FUNCTION_BLOCK Actuator2OpBase (* Composite Function Block Type *)
  (* Standard: 61499-2 *)
  (* Version 1.0.1, 9/20/2023, ApplicationLibDevTeam, Schneider Electric, First Version *)
  PACKAGE Flexbridge.FestoMPS400;
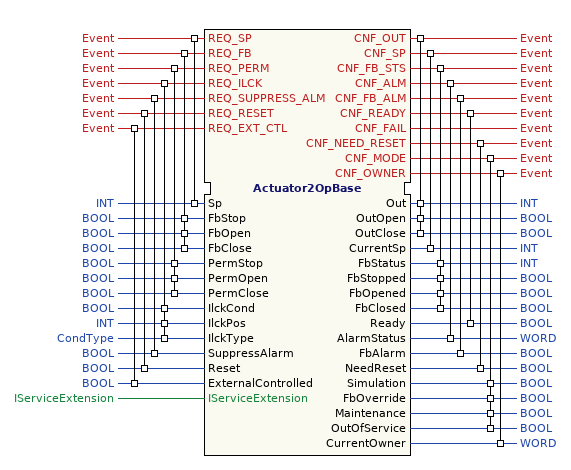
  EVENT_INPUT
    REQ_SP WITH Sp; (* Request to update setpoint *)
    REQ_FB WITH FbStop, FbOpen, FbClose; (* Request to update feedbacks *)
    REQ_PERM WITH PermStop, PermOpen, PermClose; (* Request to update permissive conditions *)
    REQ_ILCK WITH IlckCond, IlckPos, IlckType; (* Request to update interlock conditions *)
    REQ_SUPPRESS_ALM WITH SuppressAlarm; (* Request to update the alarm suppress status *)
    REQ_RESET WITH Reset; (* Request to reset the device *)
    REQ_EXT_CTL WITH ExternalControlled;
  END_EVENT
  EVENT_OUTPUT
    CNF_OUT WITH OutOpen, OutClose, Out; (* Execution confirmation of output *)
    CNF_SP WITH CurrentSp; (* Execution of confirmation Current Setpoint *)
    CNF_FB_STS WITH FbStopped, FbClosed, FbOpened, FbStatus; (* Execution of confirmed state *)
    CNF_ALM WITH AlarmStatus; (* Execution confirmation of alarm conditions *)
    CNF_FB_ALM WITH FbAlarm; (* Execution of confirmation  Fb alarm *)
    CNF_READY WITH Ready; (* Execution of Ready status *)
    CNF_FAIL; (* Execution of confirmation  failure *)
    CNF_NEED_RESET WITH NeedReset; (* Confirmation for resetting required *)
    CNF_MODE WITH Simulation, FbOverride, OutOfService, Maintenance; (* Excecution of new operational modes *)
    CNF_OWNER WITH CurrentOwner; (* Execution confirmation of owner *)
  END_EVENT
  VAR_INPUT
    Sp : INT; (* Setpoint of device (0 = Stop, 1 = Open, 2 =Close) *)
    FbStop : BOOL; (* 1 = Device stopfeedback active *)
    FbOpen : BOOL; (* 1 = Device open feedback active *)
    FbClose : BOOL; (* 1 = Device closed feedback active *)
    PermStop : BOOL := TRUE; (* 1 = Device stop permission active *)
    PermOpen : BOOL := TRUE; (* 1 = Device open permission active *)
    PermClose : BOOL := TRUE; (* 1 = Device close permission active *)
    IlckCond : BOOL; (* 1 = Interlock condition active *)
    IlckPos : INT; (* Interlock setpoint state (0 = Passive, 1 = Active1, 2 = Active2, 3 = Interlock inactive) *)
    IlckType : CondType; (* Type of condition interlock, (0 = Normal, 1 = Process interlock/Sequence interlock) *)
    SuppressAlarm : BOOL; (* 1 = Suppress alarm in HMI *)
    Reset : BOOL; (* 1 = Reset device failure *)
    ExternalControlled : BOOL; (* 1 = External control is active *)
  END_VAR
  VAR_OUTPUT
    Out : INT; (* Calculate output of the device ( 0 = Stop command, 1 = Open Command, 2 = Close Command) *)
    OutOpen : BOOL; (* 1 = Valve Output is Open *)
    OutClose : BOOL; (* 1 = Valve Output is Closed *)
    CurrentSp : INT; (* Output value considering permissive conditions *)
    FbStatus : INT; (* Confirmed state of the device (0 = Stopped, 1 = Opened, 2 = Closed,  253 = Unknown) *)
    FbStopped : BOOL; (* 1 = Stopped *)
    FbOpened : BOOL; (* 1 = Valve Open *)
    FbClosed : BOOL; (* 1 = Valve Closed *)
    Ready : BOOL; (* 1 = Device is ready to run *)
    AlarmStatus : WORD; (* Bit 1 = Device failure status, Bit 2 = Feedback failure status *)
    FbAlarm : BOOL; (* 1 = Feedback failure alarm is active *)
    NeedReset : BOOL; (* 1 = Device need reset to resume the operation *)
    Simulation : BOOL; (* 1 = Simulation mode is active *)
    FbOverride : BOOL; (* 1 = Feedback overide (Sp = FbStatus) *)
    Maintenance : BOOL; (* 1 = Maintenance mode is active *)
    OutOfService : BOOL; (* 1 = Out of service mode is active *)
    CurrentOwner : WORD; (* Current owner data from externlal source and basic owner 16#8 = Program owner, 16#10 = Operator owner, 16#4 = program Local and 16#40 Operator Local *)
  END_VAR
  SOCKETS
    IServiceExtension : IServiceExtension(ServiceState := TRUE); (* Services extension adapter(Seq control, Local panel, Maintenance and Owner) *)
  END_SOCKETS
  (* Initialization *)
  (* Supervision Interface *)
  (* Alarm Managment *)
  (* Data exchange with sequence *)
  (* Owner & Setpoint Management *)
  (* Control *)
  FBS
    plcStart : plcStart(Delay := T#0ms, Prio := 15);
    spSelection : devInSel(EnBumpless1 := FALSE, EnBumpless2 := TRUE, EnBumpless3 := FALSE, Val1 := (picosecs:=0,quality:=16#0,timestamp:=LDT#1970-01-01-05:30:00,value:=0), ResetSp := (value:=0,quality:=16#0,timestamp:=LDT#2023-01-20-10:13:38,picosecs:=0)); {SET_ATTRIBUTE(Configuration.Component.HideUnusedPorts, )}
    basicOwner : ownerControl;
    feedbackFailure : stateAlarmBasic(AlarmState := TRUE); {SET_ATTRIBUTE(HMI.AlarmText, $key:SE.App2CommonProcess.AlmLableFbFail)} {SET_ATTRIBUTE(Configuration.Component.HideUnusedPorts, )}
    progSpSelection : SELECT_24363B89CFDE21263; {SET_ATTRIBUTE(Configuration.GenericFBType.InterfaceParams, Runtime.Standard#CNT:=2;SELECT:BOOL;IN${CNT$}:INT)}
    control : valve2OpLogic(DeviceType := FALSE);
    IThis : Actuator2OpBase_HMI(QI := TRUE);
    resetConditions : DS_SELECTX_1579ED5B8ACDFC94C; {SET_ATTRIBUTE(Configuration.GenericFBType.InterfaceParams, Runtime.Standard#CNTX:=3;CNTY:=1;DI${CNTX,_,CNTY$}:BOOL)}
  END_FBS
  EVENT_CONNECTIONS
    REQ_PERM TO spSelection.REQ_SEL;
    basicOwner.CNF_OWNER TO spSelection.REQ_SEL;
    spSelection.CNF TO CNF_SP;
    REQ_FB TO control.REQ_FB;
    control.CNF_OUT TO CNF_OUT;
    control.CNF_FB_STS TO CNF_FB_STS;
    control.CNF_FB_ALM TO CNF_FB_ALM;
    control.CNF_FAIL TO CNF_FAIL;
    control.CNF_ALM TO CNF_ALM;
    control.CNF_NEED_RESET TO CNF_NEED_RESET;
    control.CNF_MODE TO CNF_MODE;
    control.CNF_READY TO CNF_READY;
    REQ_SP TO progSpSelection.REQ;
    spSelection.CNF TO IServiceExtension.CNF_STATUS;
    IServiceExtension.REQ_OWNER TO basicOwner.REQ_STDOWNER;
    REQ_SUPPRESS_ALM TO feedbackFailure.REQ_SUPRESS;
    spSelection.CNF TO control.REQ_SP;
    control.CNF_OUT TO IServiceExtension.CNF_STATUS;
    control.CNF_FB_STS TO IServiceExtension.CNF_STATUS;
    control.CNF_READY TO IServiceExtension.CNF_READY;
    REQ_PERM TO IServiceExtension.CNF_READY;
    control.CNF_NEED_RESET TO IServiceExtension.CNF_READY;
    control.CNF_ALM TO IServiceExtension.CNF_READY;
    control.CNF_ILCK TO IServiceExtension.CNF_READY;
    REQ_SUPPRESS_ALM TO IServiceExtension.CNF_SUPPRESS_ALM;
    control.CNF_MODE TO IServiceExtension.CNF_OPMODE;
    plcStart.FIRST_INIT TO IServiceExtension.CNF_SERVICE;
    feedbackFailure.INITO TO plcStart.ACK_FIRST;
    control.CNF_FB_ALM TO feedbackFailure.REQ;
    control.CNF_ILCK TO spSelection.REQ_SEL;
    IServiceExtension.REQ_CMD TO progSpSelection.REQ;
    progSpSelection.CNF TO spSelection.REQ_SP3;
    REQ_ILCK TO control.REQ_ILCK;
    REQ_EXT_CTL TO control.REQ_EXT_CTL;
    basicOwner.CNF_OWNER TO CNF_OWNER;
    REQ_RESET TO resetConditions.REQ3;
    IServiceExtension.REQ_RESET TO resetConditions.REQ2;
    resetConditions.IND TO control.REQ_RESET;
    plcStart.FIRST_INIT TO IThis.34A017503AC1070A;
    IThis.377462E9CE5193B5 TO IThis.F2953B6BB9388F21;
    feedbackFailure.CNF_ALM TO IThis.EC791CA6E67D66B3;
    spSelection.CNF TO IThis.EC791CA6E67D66B3;
    control.CNF_FB_STS TO IThis.EC791CA6E67D66B3;
    control.CNF_OUT TO IThis.EC791CA6E67D66B3;
    control.CNF_NEED_RESET TO IThis.EC791CA6E67D66B3;
    control.CNF_TRANS_FB TO IThis.EC791CA6E67D66B3;
    REQ_PERM TO IThis.EC791CA6E67D66B3;
    control.CNF_ILCK TO IThis.EC791CA6E67D66B3;
    REQ_SUPPRESS_ALM TO IThis.EC791CA6E67D66B3;
    basicOwner.CNF_OWNER TO IThis.EC791CA6E67D66B3;
    IThis.377462E9CE5193B5 TO basicOwner.REQ_BASICOWNER;
    IThis.377462E9CE5193B5 TO feedbackFailure.INIT;
    IThis.95BEA68906019444 TO control.REQ_PARA;
    IThis.95BEA68906019444 TO feedbackFailure.REQ_PARA;
    IThis.95BEA68906019444 TO IServiceExtension.CNF_CFG;
    IThis.C6CA4032A5F6989A TO spSelection.REQ_SP2;
    IThis.1A2B085F4B246BF1 TO resetConditions.REQ1;
    IThis.4711DA9A2DFC024 TO basicOwner.REQ_FORCE;
    IThis.4711DA9A2DFC024 TO control.REQ_PARA;
    IThis.4711DA9A2DFC024 TO spSelection.REQ_SEL;
    IThis.AB45C9C76752120B TO basicOwner.REQ_BASICOWNER;
  END_CONNECTIONS
  DATA_CONNECTIONS
    SuppressAlarm TO feedbackFailure.Suppress;
    PermStop TO spSelection.PermPassive;
    PermOpen TO spSelection.PermActive1;
    spSelection.PermVal TO CurrentSp;
    FbStop TO control.FbStop;
    FbOpen TO control.FbOpen;
    FbClose TO control.FbClose;
    IlckType TO control.IlckType;
    control.Out TO Out;
    control.FbStopped TO FbStopped;
    control.FbAlarm TO FbAlarm;
    control.AlarmStatus TO AlarmStatus;
    control.NeedReset TO NeedReset;
    control.Ready TO Ready;
    PermClose TO spSelection.PermActive2;
    control.FbStatus TO FbStatus;
    control.FbStatus TO IServiceExtension.Status;
    basicOwner.StdOwnerConnected TO progSpSelection.SELECT;
    Sp TO progSpSelection.IN1;
    progSpSelection.OUT TO spSelection.Val3;
    spSelection.PermVal TO IServiceExtension.CurrentSp;
    basicOwner.ProgramOwner TO spSelection.Sel3;
    basicOwner.OperatorOwner TO spSelection.Sel2;
    IServiceExtension.StdOwner TO basicOwner.StdOwner;
    spSelection.PermVal TO control.Sp;
    control.NeedReset TO IServiceExtension.NeedReset;
    control.Mode TO IServiceExtension.OpMode;
    control.Ready TO IServiceExtension.Ready;
    control.AlarmStatus TO IServiceExtension.Alarm;
    SuppressAlarm TO IServiceExtension.SuppressAlarm;
    control.Interlocked TO IServiceExtension.Interlocked;
    PermStop TO IServiceExtension.PermPassive;
    PermOpen TO IServiceExtension.PermActive1;
    PermClose TO IServiceExtension.PermActive2;
    control.FbAlarm TO feedbackFailure.Input;
    control.Interlocked TO spSelection.Ilck;
    IlckPos TO spSelection.IlckSp;
    control.Out TO IServiceExtension.CurrentOp;
    IServiceExtension.Sp TO progSpSelection.IN2;
    control.OutOpen TO OutOpen;
    control.OutClose TO OutClose;
    IlckCond TO control.IlckCond;
    control.FbOpened TO FbOpened;
    control.FbClosed TO FbClosed;
    ExternalControlled TO control.ExternalControlled;
    IlckPos TO control.IlckPos;
    basicOwner.Owner TO CurrentOwner;
    Reset TO resetConditions.DI3_1;
    IServiceExtension.Reset TO resetConditions.DI2_1;
    resetConditions.OUT1 TO control.Reset;
    control.FbStatus TO IThis.F2AD3CD6DCE76874;
    control.TransFbStatus TO IThis.18339E8B84CEF55;
    control.Out TO IThis.D2C35BC47DF71FCC;
    spSelection.PermVal TO IThis.C6876D790F3A950E;
    control.NeedReset TO IThis.9CD6749867E91606;
    basicOwner.Owner TO IThis.66F5D611520B8E21;
    feedbackFailure.AlarmStatus TO IThis.E324EF7311434CB7;
    control.Interlocked TO IThis.CAD2FBF5C8122C72;
    IlckPos TO IThis.F97E56AEBDD59492;
    PermStop TO IThis.416E212918CA047A;
    PermClose TO IThis.7DE7E04BA65FF582;
    PermOpen TO IThis.F1D46CDCC1D5A6C6;
    basicOwner.StdOwnerConnected TO IThis.9BBC553B7236462E;
    IThis.D82AC87A2FA22E86 TO basicOwner.BasicOwner;
    IThis.861B8773AF2757FC TO control.MonTime;
    IThis.5568E3E91B9AAED8 TO control.TripTime;
    IThis.3DA6D0F9276D43A4 TO control.ConfResetReq;
    IThis.4D34C1A4533BA5DF TO resetConditions.DI1_1;
    IThis.869E02415F6A841 TO spSelection.Val2;
    IThis.CF1EA84FDDBF53A1 TO Simulation;
    IThis.CF1EA84FDDBF53A1 TO control.Simulation;
    IThis.AD38F01F8F0043E7 TO FbOverride;
    IThis.AD38F01F8F0043E7 TO control.FbOverride;
    IThis.7801A8D91AA682F9 TO control.FbMode;
    IThis.C4714A0B76119976 TO OutOfService;
    IThis.C4714A0B76119976 TO spSelection.Sel1;
    IThis.C4714A0B76119976 TO control.OutOfService;
    IThis.C8DEEF765E4F14C0 TO Maintenance;
    IThis.C8DEEF765E4F14C0 TO basicOwner.ForceOperator;
    IThis.C8DEEF765E4F14C0 TO control.Maintenance;
    IThis.52A3AF601F61E85C TO spSelection.EnTrackSp;
    IThis.B394B8C6484B76DE TO feedbackFailure.ScanTime;
    IThis.E4ACFA19543211CB TO feedbackFailure.AckType;
    IThis.52A3AF601F61E85C TO IServiceExtension.EnTrackSp;
  END_CONNECTIONS
END_FUNCTION_BLOCK
